(* IEC 61131-3 sources: volt/packages/volt-lsp-iec/test-corpus/awa-palletizer/Device/Plc Logic/Application/Library Manager/L_DCO_DriveCommunication, 19 files *)

(* ---- L_DCO_COMMSTATE.dut ---- *)
TYPE L_DCO_COMMSTATE :
(
	L_DCO_STATE_BOOT := 0,
	L_DCO_STATE_INIT := 10,
	L_DCO_STATE_RESET_COMM := 20,
	L_DCO_STATE_RESET_APP := 30,
	L_DCO_STATE_PREOPERATIONAL := 40,
	L_DCO_STATE_SAVEOPERATIONAL := 50,
	L_DCO_STATE_STOPPED := 60,
	L_DCO_STATE_OPERATIONAL := 70,
	L_DCO_STATE_UNKNOWN := 80,
	L_DCO_STATE_NOT_AVAIL := 90,
	L_DCO_STATE_NOT_DETECTED := 91,
	L_DCO_STATE_NONE := 95
);
END_TYPE

(* ---- L_DCO_CONVERTDATA.dut ---- *)
TYPE L_DCO_CONVERTDATA :
UNION
	ABDATA : ARRAY [1..4] OF BYTE;
	AWDATA : ARRAY [1..2] OF WORD;
	DWDATA : DWORD;
END_UNION
END_TYPE

(* ---- L_DCO_ERROR.dut ---- *)
TYPE L_DCO_ERROR :
(
	L_DCO_NO_ERROR := 0,
	L_DCO_OTHERERROR := 20001,
	L_DCO_INVALIDINDEX := 20002,
	L_DCO_INVALIDOFFSET := 20003,
	L_DCO_INVALIDSIZE := 20004,
	L_DCO_INVALIDDATA := 20005,
	L_DCO_NOTREADY := 20006,
	L_DCO_BUSY := 20007,
	L_DCO_NOMEMORY := 20008,
	L_DCO_INVALIDPARM := 20009,
	L_DCO_INVALIDSTATE := 20010,
	L_DCO_TIMEOUT := 20011,
	L_DCO_INVALID_SLAVE_STATE := 20012,
	L_DCO_LINK_DISCONNECTED := 20013,
	L_DCO_ALL_CANNELS_BUSY := 20015,
	L_DCO_DATA_REQUEST_ERROR := 20016,
	L_DCO_BUS_OFF := 20017,
	L_DCO_SLAVE_ERROR := 20018,
	L_DCO_SDO_ABORTCODE_TOGGLE := 20020,
	L_DCO_SDO_ABORTCODE_TIMEOUT := 20021,
	L_DCO_SDO_ABORTCODE_CCS_SCS := 20022,
	L_DCO_SDO_ABORTCODE_BLK_SIZE := 20023,
	L_DCO_SDO_ABORTCODE_SEQNO := 20024,
	L_DCO_SDO_ABORTCODE_CRC := 20025,
	L_DCO_SDO_ABORTCODE_MEMORY := 20026,
	L_DCO_SDO_ABORTCODE_ACCESS := 20027,
	L_DCO_SDO_ABORTCODE_WRITEONLY := 20028,
	L_DCO_SDO_ABORTCODE_READONLY := 20029,
	L_DCO_SDO_ABORTCODE_INDEX := 20030,
	L_DCO_SDO_ABORTCODE_PDO_MAP := 20031,
	L_DCO_SDO_ABORTCODE_PDO_LEN := 20032,
	L_DCO_SDO_ABORTCODE_P_INCOMP := 20033,
	L_DCO_SDO_ABORTCODE_I_INCOMP := 20034,
	L_DCO_SDO_ABORTCODE_HARDWARE := 20035,
	L_DCO_SDO_ABORTCODE_DATA_SIZE := 20036,
	L_DCO_SDO_ABORTCODE_DATA_SIZE1 := 20037,
	L_DCO_SDO_ABORTCODE_DATA_SIZE2 := 20038,
	L_DCO_SDO_ABORTCODE_OFFSET := 20039,
	L_DCO_SDO_ABORTCODE_DATA_RANGE := 20040,
	L_DCO_SDO_ABORTCODE_DATA_RANGE1 := 20041,
	L_DCO_SDO_ABORTCODE_DATA_RANGE2 := 20042,
	L_DCO_SDO_ABORTCODE_MINMAX := 20043,
	L_DCO_SDO_ABORTCODE_GENERAL := 20044,
	L_DCO_SDO_ABORTCODE_TRANSFER := 20045,
	L_DCO_SDO_ABORTCODE_TRANSFER1 := 20046,
	L_DCO_SDO_ABORTCODE_TRANSFER2 := 20047,
	L_DCO_SDO_ABORTCODE_DICTIONARY := 20048,
	L_DCO_SDO_ABORTCODE_UNKNOWN := 20049,
	L_DCO_TRANSFERTABLE_INVALID := 20060
);
END_TYPE

(* ---- L_DCO_SDODATA.dut ---- *)
TYPE L_DCO_SDODATA :
STRUCT
	WPARAM : WORD;
	BYSUBINDEX : BYTE;
	WSTATE : WORD;
	DWOWNER : __XWORD;
	DWDATA : DWORD;
	PSDATA : POINTER TO BYTE;
	UIDATALENGTH : UINT;
	WERROR : WORD;
	WINTSTATE : WORD;
END_STRUCT
END_TYPE

(* ---- L_DCO_TRANFERDATA.dut ---- *)
TYPE L_DCO_TRANFERDATA :
STRUCT
	WINDEX : WORD;
	BYSUBINDEX : BYTE;
	DWDATA : DWORD;
	BYNROFBYTE : BYTE;
	XENABLE : BOOL;
	XWRITEACCESS : BOOL;
	XCONSIDERIDXOFFSET : BOOL;
END_STRUCT
END_TYPE

(* ---- GETBOOLEANPROPERTY.pou ---- *)
FUNCTION GETBOOLEANPROPERTY : BOOL
VAR_INPUT
	STKEY : WSTRING;
END_VAR
END_FUNCTION

(* ---- GETCOMPANY.pou ---- *)
FUNCTION GETCOMPANY : WSTRING
END_FUNCTION

(* ---- GETNUMBERPROPERTY.pou ---- *)
FUNCTION GETNUMBERPROPERTY : DINT
VAR_INPUT
	STKEY : WSTRING;
END_VAR
END_FUNCTION

(* ---- GETTEXTPROPERTY.pou ---- *)
FUNCTION GETTEXTPROPERTY : WSTRING
VAR_INPUT
	STKEY : WSTRING;
END_VAR
END_FUNCTION

(* ---- GETTEXTPROPERTY2.pou ---- *)
FUNCTION GETTEXTPROPERTY2 : POINTER TO WSTRING
VAR_INPUT
	STKEY : WSTRING;
END_VAR
END_FUNCTION

(* ---- GETTITLE.pou ---- *)
FUNCTION GETTITLE : WSTRING
END_FUNCTION

(* ---- GETVERSION.pou ---- *)
FUNCTION GETVERSION : VERSION
END_FUNCTION

(* ---- GETVERSIONPROPERTY.pou ---- *)
FUNCTION GETVERSIONPROPERTY : VERSION
VAR_INPUT
	STKEY : WSTRING;
END_VAR
END_FUNCTION

(* ---- GLOBALTEXTLIST.pou ---- *)
FUNCTION_BLOCK GLOBALTEXTLIST
VAR
	M_TEXTLISTFILE : STRING(255);
	_STNAMESPACE : STRING;
END_VAR
END_FUNCTION_BLOCK

(* ---- L_DCO_AXIS_REF_BASE.pou ---- *)
FUNCTION_BLOCK L_DCO_AXIS_REF_BASE EXTENDS IoDrvBase
VAR_INPUT
	UDITIMEOUT : UDINT := 10000;
	USICHANNEL : USINT := 1;
	ASDOREADDATA : ARRAY [1..c_wSdoMaxNumTotal] OF L_DCO_SdoData;
	ASDOWRITEDATA : ARRAY [1..c_wSdoMaxNumTotal] OF L_DCO_SdoData;
END_VAR
VAR_OUTPUT
	UIDEVICEID : UINT := 0;
	UINETID : UINT := 0;
	XCOMMUNICATIONOK : BOOL := FALSE;
	ECOMMUNICATIONSTATE : L_DCO_CommState := 0;
	AXISNAME : STRING := '';
END_VAR
VAR
	DWAXISID : DWORD;
	AXISINSTANCE : __XWORD;
	READIDX : DWORD := 1;
	WRITEIDX : DWORD := 1;
	M_PSLAVECONNECTOR : POINTER TO IoConfigConnector;
	M_PAXISCONNECTOR : POINTER TO IoConfigConnector;
	M_IIODRV : ICmpIoDrv;
	M_IIODRVPARAMETER : ICmpIoDrvParameter;
	XCOPYDATA : BOOL := TRUE;
	SINSTANCESTR : STRING;
	XPARACCESSBYSEMANOTSUPPORTED : BOOL := TRUE;
	DWSEMAPARREADACCESS : DWORD;
	DWSEMAPARWRITEACCESS : DWORD;
	C_WSDOMAXNUMTOTAL : WORD := 10;
	C_WSDOMAXNUM : WORD := 5;
	WMAXSDONUMBERREAD : WORD;
	WMAXSDONUMBERREADTOTAL : WORD;
	WMAXSDONUMBERWRITE : WORD;
	WMAXSDONUMBERWRITETOTAL : WORD;
END_VAR
END_FUNCTION_BLOCK

METHOD GETAXISSLOT : UINT
END_METHOD

METHOD GETREADPARAMETERCONTAINER : POINTER TO L_DCO_SDOData
END_METHOD

METHOD GETWRITEPARAMETERCONTAINER : POINTER TO L_DCO_SDOData
END_METHOD

METHOD INITIALIZE : UDINT
VAR_INPUT
	WMODULETYPE : UINT;
	DWINSTANCE : UDINT;
	PCONNECTOR : POINTER TO IoConfigConnector;
END_VAR
END_METHOD

METHOD IODRVREADPARAMETER : UDINT
VAR_INPUT
	PCONNECTOR : POINTER TO IoConfigConnector;
	PPARAMETER : POINTER TO IoConfigParameter;
	PDATA : POINTER TO BYTE;
	DWBITSIZE : DWORD;
	DWBITOFFSET : DWORD;
END_VAR
END_METHOD

METHOD IODRVWRITEPARAMETER : UDINT
VAR_INPUT
	PCONNECTOR : POINTER TO IoConfigConnector;
	PPARAMETER : POINTER TO IoConfigParameter;
	PDATA : POINTER TO BYTE;
	DWBITSIZE : DWORD;
	DWBITOFFSET : DWORD;
END_VAR
END_METHOD

METHOD QUERYINTERFACE : POINTER TO POINTER TO BYTE
VAR_INPUT
	IID : DWORD;
	PRESULT : POINTER TO UDINT;
END_VAR
END_METHOD

METHOD FB_INIT : BOOL
VAR_INPUT
	BINITRETAINS : BOOL;
	BINCOPYCODE : BOOL;
END_VAR
END_METHOD

(* ---- L_DCO_READDRIVEPARAMETER.pou ---- *)
FUNCTION_BLOCK L_DCO_READDRIVEPARAMETER
VAR_INPUT
	XEXECUTE : BOOL := FALSE;
	WINDEX : WORD := 0;
	BYSUBINDEX : BYTE := 0;
	XUSEINDEXASPARAM : BOOL := FALSE;
END_VAR
VAR_OUTPUT
	XDONE : BOOL := FALSE;
	XBUSY : BOOL := FALSE;
	XERROR : BOOL := FALSE;
	EERROR : L_DCO_Error := L_DCO_Error.L_DCO_No_Error;
	DWDATA : DWORD := 0;
	BYNROFBYTE : BYTE := 0;
END_VAR
VAR_IN_OUT
	AXIS : L_DCO_AXIS_REF_BASE;
END_VAR
VAR
	IDX : DWORD;
	XEXECUTEOLD : BOOL;
	SDOREAD : POINTER TO L_DCO_SdoData;
	SDOMAXREADNUM : WORD;
	SAXISNAME : STRING;
	SDOREADINTERNAL : BOOL := FALSE;
	SDONUMSTART : WORD;
	SDONUMEND : WORD;
	AXISINSTANCE : __XWORD := 0;
	XRESETOUTPUTS : BOOL;
	ABORT : BOOL;
	SDOACCESSAXISREF : BOOL;
END_VAR
END_FUNCTION_BLOCK

(* ---- L_DCO_READDRIVEPARAMETERSTRING.pou ---- *)
FUNCTION_BLOCK L_DCO_READDRIVEPARAMETERSTRING
VAR_INPUT
	XEXECUTE : BOOL := FALSE;
	WINDEX : WORD := 0;
	BYSUBINDEX : BYTE := 0;
	XUSEINDEXASPARAM : BOOL := FALSE;
END_VAR
VAR_OUTPUT
	XDONE : BOOL := FALSE;
	XBUSY : BOOL := FALSE;
	XERROR : BOOL := FALSE;
	EERROR : L_DCO_Error := L_DCO_Error.L_DCO_No_Error;
	SVALUE : STRING(255) := '';
	BYNROFBYTE : BYTE := 0;
END_VAR
VAR_IN_OUT
	AXIS : L_DCO_AXIS_REF_BASE;
END_VAR
VAR
	IDX : DWORD;
	XSEMASUPPORTEDBYAXIS : BOOL;
	XEXECUTEOLD : BOOL;
	XSEMASUPPORT : BOOL;
	SDOREAD : POINTER TO L_DCO_SdoData;
	SDONUMSTART : WORD;
	SDONUMEND : WORD;
	SDOREADINTERNAL : BOOL := FALSE;
	AXISINSTANCE : __XWORD := 0;
	SVALUEINT : STRING(255) := '';
	SAXISNAME : STRING;
	XRESETOUTPUTS : BOOL;
	ABORT : BOOL;
	SDOACCESSAXISREF : BOOL;
END_VAR
END_FUNCTION_BLOCK

(* ---- L_DCO_TRANSFERDRIVEPARAMETER.pou ---- *)
FUNCTION_BLOCK L_DCO_TRANSFERDRIVEPARAMETER
VAR_INPUT
	XEXECUTE : BOOL := FALSE;
	PSCPARAMETERDATA : POINTER TO L_DCO_TranferData;
	DWSIZEPARAMETERDATA : DWORD := 0;
	XUSEINDEXASPARAM : BOOL := FALSE;
END_VAR
VAR_OUTPUT
	XDONE : BOOL := FALSE;
	XBUSY : BOOL := FALSE;
	XERROR : BOOL := FALSE;
	EERROR : L_DCO_Error := L_DCO_Error.L_DCO_No_Error;
	WINDEXCOUNTER : WORD := 0;
END_VAR
VAR_IN_OUT
	AXIS : L_DCO_AXIS_REF_BASE;
END_VAR
VAR
	L_DCO_READDRIVEPARAMETER1 : L_DCO_ReadDriveParameter;
	L_DCO_WRITEDRIVEPARAMETER1 : L_DCO_WriteDriveParameter;
	IDX : DWORD;
	WSTEP : WORD;
	DWADRESSCOUNTER : DWORD;
	DWARRAYSIZE : DWORD;
	PSCPARAMETERDATAINTERN : POINTER TO L_DCO_TranferData;
	SCDUMMY : L_DCO_TranferData;
	DWSINGLESIZE : DWORD;
	AXISINSTANCE : __XWORD := 0;
	SAXISNAME : STRING;
END_VAR
END_FUNCTION_BLOCK

(* ---- L_DCO_WRITEDRIVEPARAMETER.pou ---- *)
FUNCTION_BLOCK L_DCO_WRITEDRIVEPARAMETER
VAR_INPUT
	XEXECUTE : BOOL := FALSE;
	WINDEX : WORD := 0;
	BYSUBINDEX : BYTE := 0;
	XUSEINDEXASPARAM : BOOL := FALSE;
	DWDATA : DWORD := 0;
	BYNROFBYTE : BYTE := 4;
END_VAR
VAR_OUTPUT
	XDONE : BOOL := FALSE;
	XBUSY : BOOL := FALSE;
	XERROR : BOOL := FALSE;
	EERROR : L_DCO_Error := L_DCO_Error.L_DCO_No_Error;
END_VAR
VAR_IN_OUT
	AXIS : L_DCO_AXIS_REF_BASE;
END_VAR
VAR
	IDX : DWORD;
	XEXECUTEOLD : BOOL;
	SDOWRITE : POINTER TO L_DCO_SdoData;
	SAXISNAME : STRING;
	SDOWRITEINTERNAL : BOOL := FALSE;
	SDONUMSTART : WORD;
	SDONUMEND : WORD;
	AXISINSTANCE : __XWORD := 0;
	XRESETOUTPUTS : BOOL;
	ABORT : BOOL;
	SDOACCESSAXISREF : BOOL;
END_VAR
END_FUNCTION_BLOCK
